Universal Robots PolyScope program: program3.urp

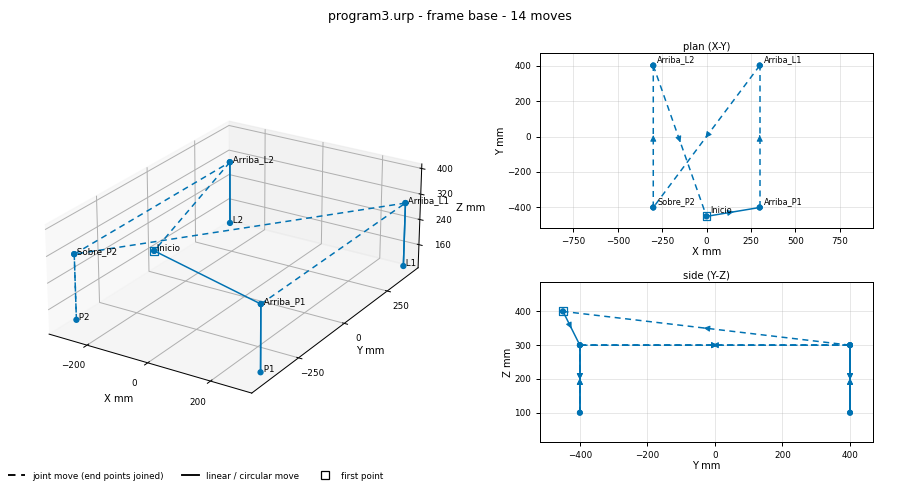
[picture p0: tool path of program3.urp in frame base, 14 of 14 moves have a stored position in this frame; points joined in program order, loops and branches not executed]
Program program3 (installation=default directory=/ursim/programs createdIn=3.15.8.106339 lastSavedIn=3.15.8.106339 robotSerialNumber=2018359999)
Calibrated DH parameters: a=[0, -0.425, -0.39225, 0, 0, 0]; d=[0.089159, 0, 0, 0.10915, 0.09465, 0.0823]; alpha=[1.570796, 0, 0, 1.570796, -1.570796, 0]; deltaTheta=[0, 0, 0, 0, 0, 0]
Robot Program (runOnlyOnce=false)
  MoveJ speed 60 deg/s, acceleration 80 deg/s^2 (useActiveTCP=true)
    Waypoint Inicio: TCP in base x=0 y=-450 z=400 mm, rx=-3.1412 ry=0 rz=0 rad; joints [75.964, -96.652, 100.886, -94.211, -90.006, 165.964] deg
  MoveL speed 250 mm/s, acceleration 1200 mm/s^2 (useActiveTCP=true) feature=Base
    Waypoint Arriba_P1: TCP in base x=300 y=-400 z=300 mm, rx=-3.1412 ry=0 rz=0 rad; joints [114.259, -86.81, 106.346, -109.514, -89.99, 204.259] deg
    Waypoint P1: TCP in base x=300 y=-400 z=100 mm, rx=-3.1412 ry=0 rz=0 rad; joints [114.259, -69.724, 120.877, -141.131, -89.99, 204.259] deg
  Set DigitalOutput (payload=1 tcpAsCog=true) pin=digital_out[1]; digitalValue=1
  Wait Sleep waitTime=0.5
  MoveL speed 250 mm/s, acceleration 1200 mm/s^2 (useActiveTCP=true) feature=Base
    Waypoint Subir_P1: TCP in base x=300 y=-400 z=300 mm, rx=-3.1412 ry=0 rz=0 rad; joints [114.259, -86.81, 106.346, -109.514, -89.99, 204.259] deg
  Wait Sleep waitTime=1
  MoveJ speed 60 deg/s, acceleration 80 deg/s^2 (useActiveTCP=true)
    Waypoint Arriba_L1: TCP in base x=300 y=400 z=300 mm, rx=-3.1412 ry=0 rz=0 rad; joints [220.518, -86.815, 106.36, -109.56, -89.982, 310.518] deg
  MoveL speed 250 mm/s, acceleration 1200 mm/s^2 (useActiveTCP=true) feature=Base
    Waypoint L1: TCP in base x=300 y=400 z=100 mm, rx=-3.1412 ry=0 rz=0 rad; joints [220.518, -69.723, 120.887, -141.18, -89.982, 310.518] deg
  Set DigitalOutput (payload=0 tcpAsCog=true) pin=digital_out[1]; digitalValue=0
  Wait Sleep waitTime=0.5
  MoveL speed 250 mm/s, acceleration 1200 mm/s^2 (useActiveTCP=true) feature=Base
    Waypoint Subir_L1: TCP in base x=300 y=400 z=300 mm, rx=-3.1412 ry=0 rz=0 rad; joints [220.518, -86.815, 106.36, -109.56, -89.982, 310.518] deg
  MoveJ speed 60 deg/s, acceleration 80 deg/s^2 (useActiveTCP=true)
    Waypoint Sobre_P2: TCP in base x=-300.017 y=-399.967 z=299.974 mm, rx=-3.1411 ry=0 rz=-0.0001 rad; joints [40.52, -86.81, 106.35, -109.52, -90.02, 130.52] deg
  MoveJ speed 60 deg/s, acceleration 80 deg/s^2 (useActiveTCP=true)
    Waypoint P2: TCP in base x=-300.016 y=-399.965 z=99.957 mm, rx=-3.1411 ry=0 rz=-0.0001 rad; joints [40.52, -69.72, 120.88, -141.14, -90.02, 130.52] deg
  Set DigitalOutput (payload=1 tcpAsCog=true) pin=digital_out[1]; digitalValue=1
  Wait Sleep waitTime=0.5
  MoveJ speed 60 deg/s, acceleration 80 deg/s^2 (useActiveTCP=true)
    Waypoint Subir_P2: TCP in base x=-300.017 y=-399.967 z=299.974 mm, rx=-3.1411 ry=0 rz=-0.0001 rad; joints [40.52, -86.81, 106.35, -109.52, -90.02, 130.52] deg
  Wait Sleep waitTime=1
  MoveJ speed 60 deg/s, acceleration 80 deg/s^2 (useActiveTCP=true)
    Waypoint Arriba_L2: TCP in base x=-299.959 y=399.993 z=300.008 mm, rx=3.1415 ry=0 rz=0.0007 rad; joints [-65.74, -86.814, 106.35, -109.52, -90.02, 24.26] deg
  MoveL speed 250 mm/s, acceleration 1200 mm/s^2 (useActiveTCP=true) feature=Base
    Waypoint L2: TCP in base x=-299.964 y=400.004 z=99.95 mm, rx=3.1414 ry=0 rz=0.0007 rad; joints [-65.74, -69.719, 120.88, -141.14, -90.02, 24.26] deg
  Set DigitalOutput (payload=0 tcpAsCog=true) pin=digital_out[1]; digitalValue=0
  Wait Sleep waitTime=0.5
  MoveL speed 250 mm/s, acceleration 1200 mm/s^2 (useActiveTCP=true) feature=Base
    Waypoint Subir_L2: TCP in base x=-299.959 y=399.993 z=300.008 mm, rx=3.1415 ry=0 rz=0.0007 rad; joints [-65.74, -86.814, 106.35, -109.52, -90.02, 24.26] deg
  MoveJ speed 60 deg/s, acceleration 80 deg/s^2 (useActiveTCP=true)
    Waypoint Fin: TCP in base x=0 y=-450 z=400 mm, rx=-3.1412 ry=0 rz=0 rad; joints [75.964, -96.652, 100.886, -94.211, -90.006, 165.964] deg
  Wait DigitalInput pin=digital_in[0]; digitalValue=1
